(* IEC 61131-3 sources: RootPLC/conformance/cases/diff, 4 files *)

(* ---- ok_diff_adapter_agrees.st ---- *)
(* spec: [diff.command] [diff.interface] [diff.stimuli] [diff.compare] [diff.report] [diff.limits]
   expect: ok *)
(* A reference start/stop latch and a block written another way, with
   other names, wrapped in an adapter that has the reference's names.
   rootplc diff --reference FB_RefLatch --unit FB_LatchAdapter agrees
   (crates/rootplc-driver/tests/diff.rs). *)
FUNCTION_BLOCK FB_RefLatch
VAR_INPUT
    Start  : BOOL;
    StopOk : BOOL;                 (* FALSE stops; stop wins *)
    Limit  : REAL;
    Level  : REAL;
END_VAR
VAR_OUTPUT
    Out  : BOOL;
    High : BOOL;                   (* Level above Limit *)
END_VAR
IF NOT StopOk THEN
    Out := FALSE;
ELSIF Start THEN
    Out := TRUE;
END_IF;
High := Level > Limit;
END_FUNCTION_BLOCK

(* the block from a real project: other names, other style *)
FUNCTION_BLOCK FB_PumpLatch
VAR_INPUT
    xStart     : BOOL;
    xStopNC    : BOOL;
    rThreshold : REAL;
    rValue     : REAL;
END_VAR
VAR_OUTPUT
    xRun   : BOOL;
    xAlarm : BOOL;
END_VAR
VAR
    latch : RS;
END_VAR
latch(S := xStart, R1 := NOT xStopNC);
xRun := latch.Q1;
xAlarm := NOT (rValue <= rThreshold);
END_FUNCTION_BLOCK

(* the adapter: the reference's names around the real block *)
FUNCTION_BLOCK FB_LatchAdapter
VAR_INPUT
    Start  : BOOL;
    StopOk : BOOL;
    Limit  : REAL;
    Level  : REAL;
END_VAR
VAR_OUTPUT
    Out  : BOOL;
    High : BOOL;
END_VAR
VAR
    wrapped : FB_PumpLatch;
END_VAR
wrapped(xStart := Start, xStopNC := StopOk, rThreshold := Limit, rValue := Level);
Out := wrapped.xRun;
High := wrapped.xAlarm;
END_FUNCTION_BLOCK

(* ---- ok_diff_finds_a_difference.st ---- *)
(* spec: [diff.compare] [diff.report] [diff.stimuli]
   expect: ok *)
(* A latch where start wins over stop, compared with a reference where stop
   wins: rootplc diff --reference FB_StopWins --unit FB_StartWins reports a
   difference on Out in the cycle where Start and a stop come together
   (crates/rootplc-driver/tests/diff.rs). With --set StopOk=TRUE the
   difference cannot occur and the blocks agree. *)
FUNCTION_BLOCK FB_StopWins
VAR_INPUT
    Start  : BOOL;
    StopOk : BOOL;
    Delay  : TIME := T#1s;
END_VAR
VAR_OUTPUT
    Out   : BOOL;
    Since : TIME;
END_VAR
VAR
    t : TON;
END_VAR
IF NOT StopOk THEN
    Out := FALSE;
ELSIF Start THEN
    Out := TRUE;
END_IF;
t(IN := Out, PT := Delay);
Since := t.ET;
END_FUNCTION_BLOCK

FUNCTION_BLOCK FB_StartWins
VAR_INPUT
    Start  : BOOL;
    StopOk : BOOL;
    Delay  : TIME := T#1s;
END_VAR
VAR_OUTPUT
    Out   : BOOL;
    Since : TIME;
END_VAR
VAR
    t : TON;
END_VAR
IF Start THEN
    Out := TRUE;
ELSIF NOT StopOk THEN
    Out := FALSE;
END_IF;
t(IN := Out, PT := Delay);
Since := t.ET;
END_FUNCTION_BLOCK

(* ---- ok_diff_slice.st ---- *)
(* spec: [diff.slice]
   expect: ok *)
(* A unit that uses a type and a helper block declared elsewhere in the
   project. rootplc diff keeps the files that declare FB_Ref, FB_Uses and
   what they use (here all in this file); a broken file of the same project
   that neither block needs is left out
   (crates/rootplc-driver/tests/diff.rs). *)
TYPE E_Level : (Low, High); END_TYPE

FUNCTION_BLOCK FB_Helper
VAR_INPUT x : REAL; END_VAR
VAR_OUTPUT level : E_Level; END_VAR
IF x > 50.0 THEN
    level := E_Level#High;
ELSE
    level := E_Level#Low;
END_IF;
END_FUNCTION_BLOCK

FUNCTION_BLOCK FB_Ref
VAR_INPUT x : REAL; END_VAR
VAR_OUTPUT high : BOOL; END_VAR
high := x > 50.0;
END_FUNCTION_BLOCK

FUNCTION_BLOCK FB_Uses
VAR_INPUT x : REAL; END_VAR
VAR_OUTPUT high : BOOL; END_VAR
VAR h : FB_Helper; END_VAR
h(x := x);
high := h.level = E_Level#High;
END_FUNCTION_BLOCK

(* ---- warn_whitebox_adapter.st ---- *)
(* spec: [diff.adapter] [tests.whitebox]
   expect: warning RP0136
   run: PRG_Main cycles=2
   assert: out = TRUE *)
(* A device block that keeps its I/O internal (mapped AT %I* in a vendor
   tool), and a white-box adapter that drives it through its internal
   variables, as rootplc diff needs. *)
FUNCTION_BLOCK FB_Device
VAR
    sensor : BOOL;
    coil   : BOOL;
END_VAR
coil := sensor;
END_FUNCTION_BLOCK

{attribute 'rootplc.adapter'}
FUNCTION_BLOCK FB_DeviceAdapter
VAR_INPUT
    In : BOOL;
END_VAR
VAR_OUTPUT
    Out : BOOL;
END_VAR
VAR
    dev : FB_Device;
END_VAR
dev.sensor := In;
dev();
Out := dev.coil;
END_FUNCTION_BLOCK

PROGRAM PRG_Main
VAR
    a   : FB_DeviceAdapter;
    out : BOOL;
END_VAR
a(In := TRUE);
out := a.Out;
END_PROGRAM
